Fanuc KAREL source: kc00018.KL

-- PROVISIONAL review KL for V770-1; original PC SHA256 7015e8e1d003445605343b9f4293a88e8323d26ab47f5b3b7ab9f676c812802e
-- Incomplete behavior may be omitted. Consult companion uncertainty JSON. Do not deploy.
PROGRAM KC00018
%NOLOCKGROUP
BEGIN
  -- UNRESOLVED_PC offsets 5-63; opcodes 27,22,2A,22,2A,22,22,2A,22,22,22,22,31
  -- UNRESOLVED_PC offsets 68-72; opcodes 7F
END KC00018
